FUNCTION_BLOCK fbBistableDoubleCoilRelay IMPLEMENTS iRelay
VAR_OUTPUT
	RelaySetOutput AT %Q* : BOOL;
	RelayResetOutput AT %Q* : BOOL;
END_VAR
VAR
	CmdSet : BOOL;
    CmdReset : BOOL;
    SetPulseTP : TP;
    ResetPulseTP : TP;
END_VAR
VAR CONSTANT
    PulseTime : TIME := T#200MS;
END_VAR
VAR RETAIN
	RelaySet : BOOL;
END_VAR

// Interlock commands
IF CmdReset THEN
	CmdSet := FALSE;
	RelaySet := FALSE;
ELSIF CmdSet THEN
	CmdReset := FALSE;
	RelaySet := TRUE;
END_IF


SetPulseTP(IN := CmdSet, PT := PulseTime);
ResetPulseTP(IN := CmdReset, PT := PulseTime);

// Pulse physical outputs
RelaySetOutput := SetPulseTP.Q;
RelayResetOutput := ResetPulseTP.Q;

// Reset commands
CmdSet := FALSE;
CmdReset := FALSE;

{warning 'Add property implementation'}
PROPERTY IsSet : BOOL
GET
IsSet := RelaySet;
END_GET
END_PROPERTY

{warning 'Add method implementation '}
METHOD Reset
CmdReset := TRUE;
END_METHOD

{warning 'Add method implementation '}
METHOD Set
CmdSet := TRUE;
END_METHOD

END_FUNCTION_BLOCK

(* stored: Version 1.1.0.1
   POU fbBistableDoubleCoilRelay: Id {335a84c2-d420-4524-aa4e-8efe9b956cf1}, SpecialFunc None
   Property IsSet: Id {c31de52c-601a-4de2-9ac8-9f8bfedf0563}
   Get Get: Id {9d09fda1-2f39-4c3c-8790-750d752761be}
   Method Reset: Id {cad43598-7528-4a0d-9bc6-4e05f8803093}
   Method Set: Id {276ef09e-4879-413f-bd8a-3a7e49269787} *)
